FUNCTION_BLOCK FB_StartGame
VAR_INPUT
END_VAR
VAR_OUTPUT
END_VAR
VAR
END_VAR

END_FUNCTION_BLOCK

(* stored: Version 1.1.0.1, ProductVersion 3.1.4024.15
   POU FB_StartGame: Id {a2e1a3e2-4725-41ee-97fe-88b1fce1b3a5}, SpecialFunc None *)
